Fanuc KAREL source: KT00179.KL

PROGRAM KT00179
%NOLOCKGROUP
VAR
  Y1: ARRAY[2] OF BYTE
  R2: REAL
  OUT: INTEGER
BEGIN
  Y1[1] = 2
    R2 = 3.0
  OUT = Y1[1] MOD R2
END KT00179
